// TIA Portal V21 export
// export: Created 2026-11-08T21:35:43.7186227Z, ExportSetting WithDefaults, DisplayName Totally Integrated Automation Portal, DisplayVersion V21 Update 3, DisplayName STEP 7 Professional, DisplayVersion V21 Update 3, DisplayName STEP 7 Safety, DisplayVersion V21, DisplayName Tech WebApplication, DisplayVersion V21, DisplayName WinCC Basic/Comfort/Advanced, DisplayVersion V21 Update 3, DisplayName WinCC Unified, DisplayVersion V21 Update 3
FUNCTION_BLOCK "FB_StlC_055"   // FB79, STL
TITLE = STL call BLKMOV
{ S7_Optimized_Access := 'FALSE' }
VERSION : 0.1
// stored: AutoNumber true, UDAEnableTagReadback false
   VAR_OUTPUT
      io : Int;
   END_VAR
BEGIN

NETWORK
TITLE = 055 BLKMOV
      CALL  BLKMOV
      ( SRCBLK  := "DB_Arr"."a",
        RET_VAL := #io,
        DSTBLK  := "DB_Arr"."b"
      );

NETWORK
TITLE = 056 UBLKMOV
      CALL  UBLKMOV
      ( SRCBLK  := "DB_Arr"."a",
        RET_VAL := #io,
        DSTBLK  := "DB_Arr"."b"
      );
END_FUNCTION_BLOCK
